Fanuc KAREL source: kx00014.KL

PROGRAM KX00014
%STACKSIZE=65535
%PRIORITY=65535
%NOLOCKGROUP
VAR
I : INTEGER
J : INTEGER
B : BOOLEAN
F : FILE
S : STRING[80]
P : XYZWPR
BEGIN
-- UNRESOLVED_PC line 11 opcodes [9D 3C] marker_code=0
END KX00014
